// Current language of the event texts.
INTERFACE I_LanguageProvider

PROPERTY Current : E_Language
GET
END_GET
END_PROPERTY

END_INTERFACE

(* stored: Version 1.1.0.1, ProductVersion 3.1.4026.26
   Itf I_LanguageProvider: Id {2d129caa-51c4-4106-a1db-be6b4dfcc74e}
   Property Current: Id {62175160-0d42-4ab2-b8e7-0f8ae29f5978}
   Get Get: Id {6edbf9ee-113b-46a8-b495-0296f87a9f11} *)
